// TwinCAT 3 PLC project PLC
// ProgramVersion: 3.1.4026.26
// libraries:
//   Tc2_Standard, * (Beckhoff Automation GmbH)
//   Tc2_System, * (Beckhoff Automation GmbH)
//   Tc3_IotBase, * (Beckhoff Automation GmbH)
// project tree:
//   FBs/ FB_BenchMqttEcho.TcPOU
//   GVLs/ GVL.TcGVL, GVL_Bench.TcGVL
//   / PlcTask.TcTTO
//   POUs/ MAIN.TcPOU, PRG_Echo.TcPOU, PRG_EchoMqtt.TcPOU

CONFIGURATION PLC
    RESOURCE PLC ON TwinCAT3
        TASK PlcTask(INTERVAL := T#1ms, PRIORITY := 20);
        PROGRAM MAIN WITH PlcTask : MAIN;
    END_RESOURCE
END_CONFIGURATION

// ---- GVLs/GVL.TcGVL
// Áreas do servidor Modbus TCP (TF6250), a partir do endereço 32768.
// Sem 'qualified_only': o servidor Modbus procura estas variáveis pelo nome.
VAR_GLOBAL
    mb_Input_Coils      : ARRAY [0..255] OF BOOL;
    mb_Output_Coils     : ARRAY [0..255] OF BOOL;
    mb_Input_Registers  : ARRAY [0..255] OF WORD;
    mb_Output_Registers : ARRAY [0..255] OF WORD;
END_VAR

// ---- GVLs/GVL_Bench.TcGVL
{attribute 'qualified_only'}
VAR_GLOBAL
    {attribute 'OPC.UA.DA' := '1'}
    nIn  : DINT;   // escrito pelo cliente (Python)
    {attribute 'OPC.UA.DA' := '1'}
    nOut : DINT;   // eco: PRG_Echo copia nIn aqui a cada ciclo
END_VAR

// ---- POUs/MAIN.TcPOU
PROGRAM MAIN
VAR
END_VAR

PRG_Echo();
PRG_EchoMqtt();

END_PROGRAM

// ---- POUs/PRG_Echo.TcPOU
PROGRAM PRG_Echo
VAR
END_VAR

// Eco usado pelo benchmark: devolve, no mesmo ciclo, o que o cliente escreveu.
// ADS e OPC UA: DINT.
GVL_Bench.nOut := GVL_Bench.nIn;

// Modbus TCP: o cliente escreve o holding register (função 6) e lê o input register (função 4).
GVL.mb_Input_Registers[0] := GVL.mb_Output_Registers[0];

END_PROGRAM

// ---- POUs/PRG_EchoMqtt.TcPOU
(*
    Chama o eco MQTT. É um programa à parte do PRG_Echo de propósito: usar o MQTT exige a
    TF6701 e a referência Tc3_IotBase; quem só mede ADS, OPC UA e Modbus não precisa disso.
    Para medir MQTT: importe FB_BenchMqttEcho e este programa, adicione a referência
    Tc3_IotBase, ajuste o endereço do broker abaixo e chame PRG_EchoMqtt() no MAIN.
*)
PROGRAM PRG_EchoMqtt
VAR
    fbEcho : FB_BenchMqttEcho;
    xHabilita : BOOL := TRUE; // pode ser forçado a FALSE para desconectar
END_VAR

fbEcho(bEnable   := xHabilita,
       sHost     := '10.199.162.30',   // o mesmo broker de [mqtt] host no config.toml
       nPort     := 1883,
       sTopicIn  := 'bench/in',
       sTopicOut := 'bench/out');

END_PROGRAM

// ---- FBs/FB_BenchMqttEcho.TcPOU
(*
    Eco MQTT do benchmark: assina sTopicIn e devolve, em sTopicOut, o mesmo payload.

    Exige a TF6701 (IoT Communication MQTT) e a referência Tc3_IotBase no projeto PLC.
    A conexão, a fila de entrada (ipMessageQueue), o Subscribe e o Dequeue seguem o
    FB_DfiMqttSubscriber do projeto CX9240_DataFlowInventory, validado em bancada. O que
    este FB acrescenta é o Publish, conferido apenas na documentação da Beckhoff (TF6701,
    FB_IotMqttClient.Publish) e AINDA NÃO TESTADO no XAE.

    Uma mensagem por ciclo (mesma contrapressão do DrainOneMessage do DFI).
    O payload é texto ASCII (o número em decimal) e volta sem alteração.
*)
FUNCTION_BLOCK FB_BenchMqttEcho
VAR_INPUT
    bEnable   : BOOL;
    sHost     : STRING(80) := '192.168.1.10'; // broker
    nPort     : UINT := 1883;
    sTopicIn  : STRING(80) := 'bench/in';
    sTopicOut : STRING(80) := 'bench/out';
END_VAR
VAR_OUTPUT
    bConnected : BOOL;
    bError     : BOOL;
    nEchoed    : UDINT; // mensagens devolvidas
END_VAR
VAR
    fbMqtt        : FB_IotMqttClient;
    fbMsgQueue    : Tc3_IotBase.FB_IotMqttMessageQueue; // fila de entrada: o client não a cria sozinho
    fbMessage     : Tc3_IotBase.FB_IotMqttMessage;
    bParamsSet    : BOOL;
    bSubscribed   : BOOL;
    bWasConnected : BOOL;
    sTopicSub     : STRING(80); // Subscribe e Publish recebem o tópico por referência
    sTopicPub     : STRING(80);
    sPayload      : STRING(63);
END_VAR

// -- desabilitado: derruba a conexão e zera o handshake de assinatura --
IF NOT bEnable THEN
    fbMqtt.Execute(bConnect := FALSE);
    bConnected    := FALSE;
    bSubscribed   := FALSE;
    bWasConnected := FALSE;
    RETURN;
END_IF

// -- parametrização única (igual ao ApplyBrokerParams do DFI) --
IF NOT bParamsSet THEN
    fbMqtt.sHostName      := sHost;
    fbMqtt.nHostPort      := nPort;
    fbMqtt.sClientId      := 'bench-plc-echo';
    fbMqtt.ipMessageQueue := fbMsgQueue; // sem isso a fila de entrada fica 0 para sempre
    bParamsSet := TRUE;
END_IF

// -- conexão cíclica --
fbMqtt.Execute(bConnect := TRUE);
bConnected := fbMqtt.bConnected;
bError     := fbMqtt.bError;

// a queda invalida a assinatura
IF bWasConnected AND NOT bConnected THEN
    bSubscribed := FALSE;
END_IF
bWasConnected := bConnected;

IF bConnected AND NOT bSubscribed THEN
    sTopicSub   := sTopicIn;
    bSubscribed := fbMqtt.Subscribe(sTopic := sTopicSub,
                                    eQoS   := Tc3_IotBase.TcIotMqttQos.AtLeastOnceDelivery);
END_IF

// -- eco: tira no máximo UMA mensagem por ciclo e a devolve --
IF bConnected AND bSubscribed AND (fbMsgQueue.nQueuedMessages > 0) THEN
    IF fbMsgQueue.Dequeue(fbMessage := fbMessage) THEN
        fbMessage.GetPayload(pPayload            := ADR(sPayload),
                             nPayloadSize        := SIZEOF(sPayload) - 1,
                             bSetNullTermination := TRUE);
        sTopicPub := sTopicOut;
        IF fbMqtt.Publish(sTopic       := sTopicPub,
                          pPayload     := ADR(sPayload),
                          nPayloadSize := INT_TO_UDINT(LEN(sPayload)), // sem o byte nulo: o cliente lê texto
                          eQoS         := Tc3_IotBase.TcIotMqttQos.AtLeastOnceDelivery,
                          bRetain      := FALSE,
                          bQueue       := FALSE) THEN // bQueue é reservado: sempre FALSE
            nEchoed := nEchoed + 1;
        END_IF
    END_IF
END_IF

END_FUNCTION_BLOCK
